Fanuc KAREL source: kt00649.KL

-- PROVISIONAL review KL for V1013-1; original PC SHA256 190244943c37dca6fd7ca82894e824f829b85f1d3598727c5e2f902220a74c9e
-- Incomplete behavior may be omitted. Consult companion uncertainty JSON. Do not deploy.
PROGRAM KT00649
%NOLOCKGROUP
VAR
  OUT : INTEGER
-- UNRESOLVED_DECL H1 type=002017
-- UNRESOLVED_DECL H2 type=002017
BEGIN
  -- UNRESOLVED_PC offsets 5-19; opcodes 2E,22,9D,33,B4
  -- UNRESOLVED_PC offsets 24-38; opcodes 2E,22,9D,33,B4
  -- UNRESOLVED_PC offsets 43-57; opcodes 2E,22,9D,33,B4
  -- UNRESOLVED_PC offsets 62-76; opcodes 2E,22,9D,33,B4
  -- UNRESOLVED_PC offsets 81-97; opcodes 22,9D,33,B3,51,23
  -- UNRESOLVED_PC offsets 102-106; opcodes 7F
END KT00649
